TYPE ST_StateDevice_HMI_Status :
STRUCT
	cfgDeviceName		: STRING;
	stsAuto				: BOOL;
	stsIdle				: BOOL;
	stsDone				: BOOL;
	stsRunning 			: BOOL;
	stsFaulted			: BOOL;
	stsAborting			: BOOL;
	stsAborted			: BOOL;
	stsFaultDescription	: STRING;
	stsState			: STRING;
	stsStepDescription	: STRING;
	stsStepNumber		: INT;
	stsRetryAllowed		: BOOL;
END_STRUCT
END_TYPE

(* stored: Version 1.1.0.1
   DUT ST_StateDevice_HMI_Status: Id {bf497164-7e14-4451-bf9a-5b0043fa1ae0} *)
